// TIA Portal V20 export
ORGANIZATION_BLOCK "T4_Ciclo"   // OB127, LAD, ProgramCycle
TITLE = T4_Ciclo
{ S7_Optimized_Access := 'TRUE' }
AUTHOR : IA
FAMILY : PRUEBA
VERSION : 0.1
// Tanda 1: llama a todas las pruebas
// stored: AutoNumber false, IsIECCheckEnabled false, SetENOAutomatically false
   VAR_INPUT
      Initial_Call : Bool;
      Remanence : Bool;
   END_VAR
BEGIN

REGION Network 1: T4_Base
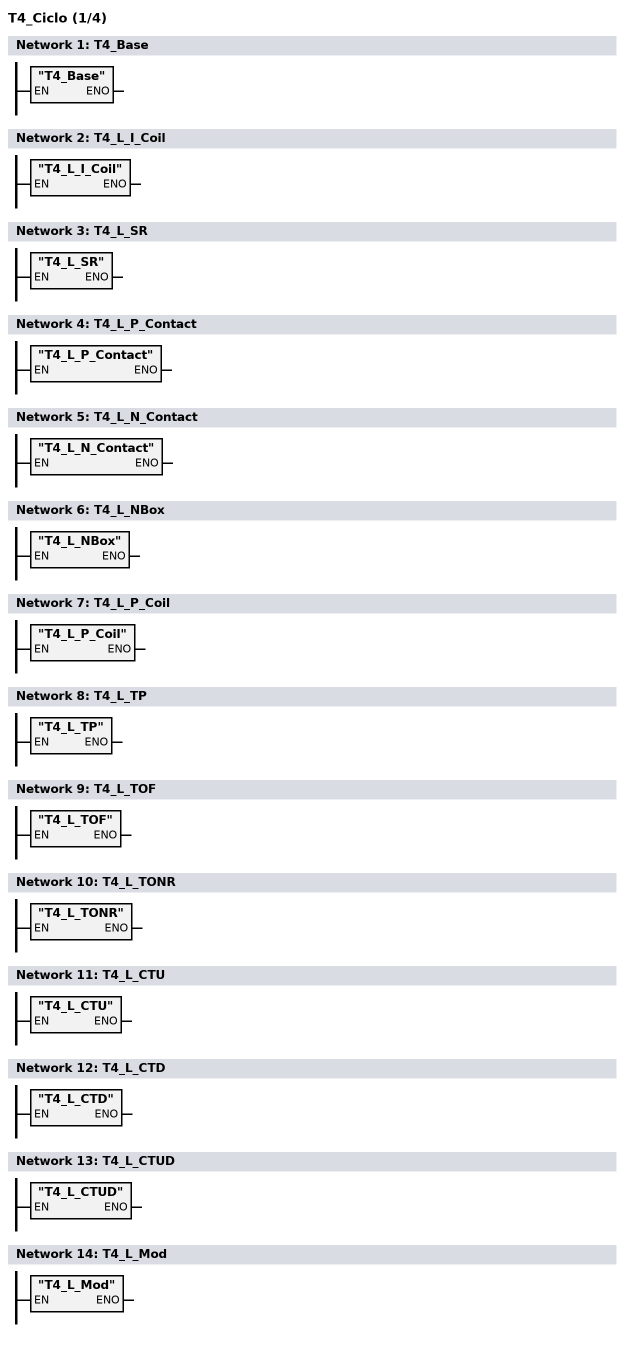
   RUNG wire#powerrail
      "T4_Base"()
   END_RUNG
   // the same network as SCL:
   "T4_Base"();
END_REGION

REGION Network 2: T4_L_I_Coil
   RUNG wire#powerrail
      "T4_L_I_Coil"()
   END_RUNG
   // the same network as SCL:
   "T4_L_I_Coil"();
END_REGION

REGION Network 3: T4_L_SR
   RUNG wire#powerrail
      "T4_L_SR"()
   END_RUNG
   // the same network as SCL:
   "T4_L_SR"();
END_REGION

REGION Network 4: T4_L_P_Contact
   RUNG wire#powerrail
      "T4_L_P_Contact"()
   END_RUNG
   // the same network as SCL:
   "T4_L_P_Contact"();
END_REGION

REGION Network 5: T4_L_N_Contact
   RUNG wire#powerrail
      "T4_L_N_Contact"()
   END_RUNG
   // the same network as SCL:
   "T4_L_N_Contact"();
END_REGION

REGION Network 6: T4_L_NBox
   RUNG wire#powerrail
      "T4_L_NBox"()
   END_RUNG
   // the same network as SCL:
   "T4_L_NBox"();
END_REGION

REGION Network 7: T4_L_P_Coil
   RUNG wire#powerrail
      "T4_L_P_Coil"()
   END_RUNG
   // the same network as SCL:
   "T4_L_P_Coil"();
END_REGION

REGION Network 8: T4_L_TP
   RUNG wire#powerrail
      "T4_L_TP"()
   END_RUNG
   // the same network as SCL:
   "T4_L_TP"();
END_REGION

REGION Network 9: T4_L_TOF
   RUNG wire#powerrail
      "T4_L_TOF"()
   END_RUNG
   // the same network as SCL:
   "T4_L_TOF"();
END_REGION

REGION Network 10: T4_L_TONR
   RUNG wire#powerrail
      "T4_L_TONR"()
   END_RUNG
   // the same network as SCL:
   "T4_L_TONR"();
END_REGION

REGION Network 11: T4_L_CTU
   RUNG wire#powerrail
      "T4_L_CTU"()
   END_RUNG
   // the same network as SCL:
   "T4_L_CTU"();
END_REGION

REGION Network 12: T4_L_CTD
   RUNG wire#powerrail
      "T4_L_CTD"()
   END_RUNG
   // the same network as SCL:
   "T4_L_CTD"();
END_REGION

REGION Network 13: T4_L_CTUD
   RUNG wire#powerrail
      "T4_L_CTUD"()
   END_RUNG
   // the same network as SCL:
   "T4_L_CTUD"();
END_REGION

REGION Network 14: T4_L_Mod
   RUNG wire#powerrail
      "T4_L_Mod"()
   END_RUNG
   // the same network as SCL:
   "T4_L_Mod"();
END_REGION

REGION Network 15: T4_L_Neg
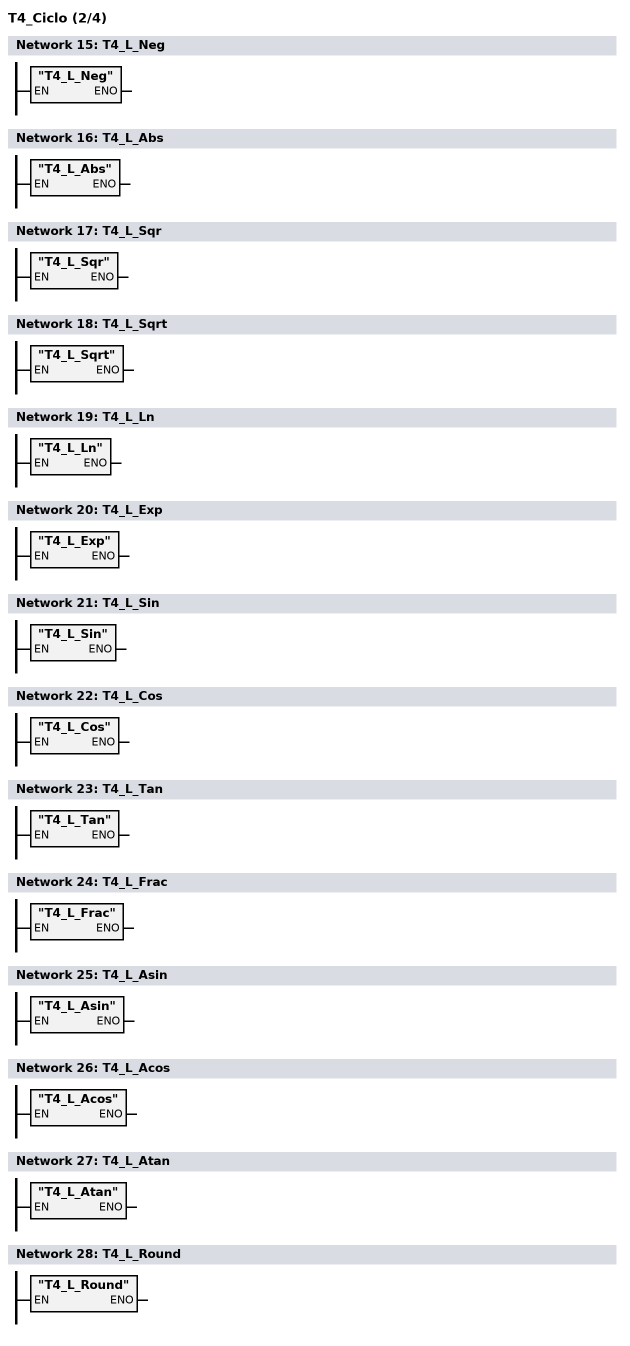
   RUNG wire#powerrail
      "T4_L_Neg"()
   END_RUNG
   // the same network as SCL:
   "T4_L_Neg"();
END_REGION

REGION Network 16: T4_L_Abs
   RUNG wire#powerrail
      "T4_L_Abs"()
   END_RUNG
   // the same network as SCL:
   "T4_L_Abs"();
END_REGION

REGION Network 17: T4_L_Sqr
   RUNG wire#powerrail
      "T4_L_Sqr"()
   END_RUNG
   // the same network as SCL:
   "T4_L_Sqr"();
END_REGION

REGION Network 18: T4_L_Sqrt
   RUNG wire#powerrail
      "T4_L_Sqrt"()
   END_RUNG
   // the same network as SCL:
   "T4_L_Sqrt"();
END_REGION

REGION Network 19: T4_L_Ln
   RUNG wire#powerrail
      "T4_L_Ln"()
   END_RUNG
   // the same network as SCL:
   "T4_L_Ln"();
END_REGION

REGION Network 20: T4_L_Exp
   RUNG wire#powerrail
      "T4_L_Exp"()
   END_RUNG
   // the same network as SCL:
   "T4_L_Exp"();
END_REGION

REGION Network 21: T4_L_Sin
   RUNG wire#powerrail
      "T4_L_Sin"()
   END_RUNG
   // the same network as SCL:
   "T4_L_Sin"();
END_REGION

REGION Network 22: T4_L_Cos
   RUNG wire#powerrail
      "T4_L_Cos"()
   END_RUNG
   // the same network as SCL:
   "T4_L_Cos"();
END_REGION

REGION Network 23: T4_L_Tan
   RUNG wire#powerrail
      "T4_L_Tan"()
   END_RUNG
   // the same network as SCL:
   "T4_L_Tan"();
END_REGION

REGION Network 24: T4_L_Frac
   RUNG wire#powerrail
      "T4_L_Frac"()
   END_RUNG
   // the same network as SCL:
   "T4_L_Frac"();
END_REGION

REGION Network 25: T4_L_Asin
   RUNG wire#powerrail
      "T4_L_Asin"()
   END_RUNG
   // the same network as SCL:
   "T4_L_Asin"();
END_REGION

REGION Network 26: T4_L_Acos
   RUNG wire#powerrail
      "T4_L_Acos"()
   END_RUNG
   // the same network as SCL:
   "T4_L_Acos"();
END_REGION

REGION Network 27: T4_L_Atan
   RUNG wire#powerrail
      "T4_L_Atan"()
   END_RUNG
   // the same network as SCL:
   "T4_L_Atan"();
END_REGION

REGION Network 28: T4_L_Round
   RUNG wire#powerrail
      "T4_L_Round"()
   END_RUNG
   // the same network as SCL:
   "T4_L_Round"();
END_REGION

REGION Network 29: T4_L_Ceil
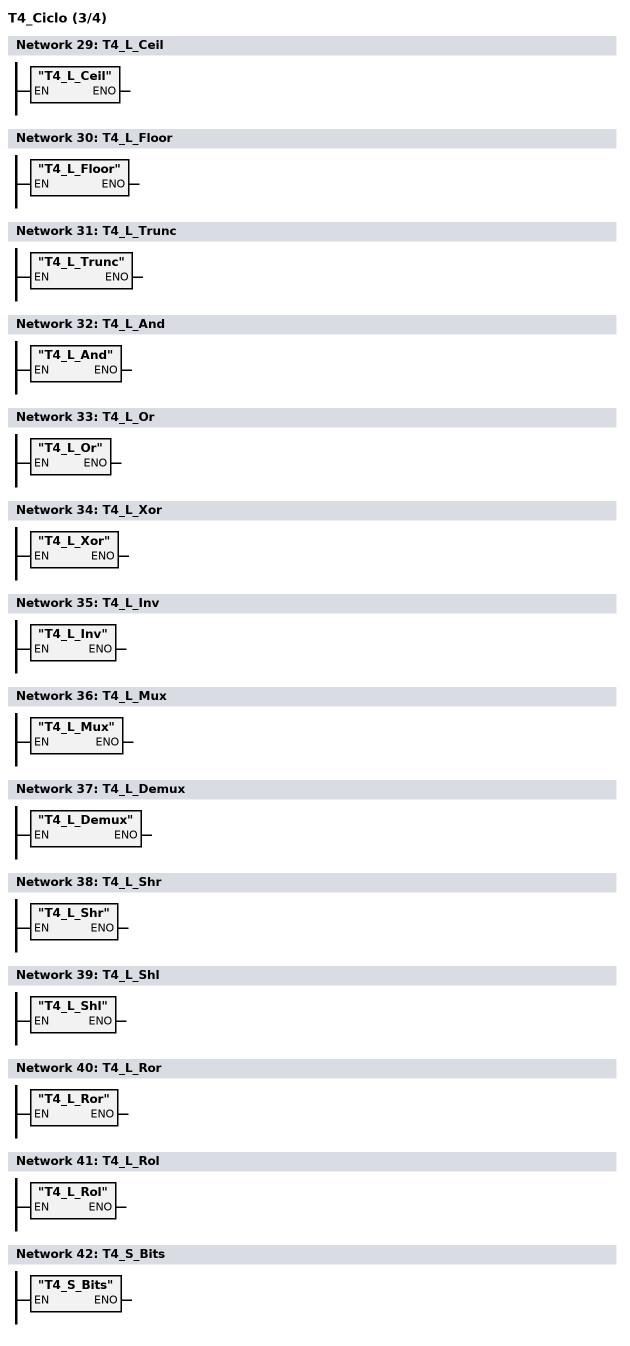
   RUNG wire#powerrail
      "T4_L_Ceil"()
   END_RUNG
   // the same network as SCL:
   "T4_L_Ceil"();
END_REGION

REGION Network 30: T4_L_Floor
   RUNG wire#powerrail
      "T4_L_Floor"()
   END_RUNG
   // the same network as SCL:
   "T4_L_Floor"();
END_REGION

REGION Network 31: T4_L_Trunc
   RUNG wire#powerrail
      "T4_L_Trunc"()
   END_RUNG
   // the same network as SCL:
   "T4_L_Trunc"();
END_REGION

REGION Network 32: T4_L_And
   RUNG wire#powerrail
      "T4_L_And"()
   END_RUNG
   // the same network as SCL:
   "T4_L_And"();
END_REGION

REGION Network 33: T4_L_Or
   RUNG wire#powerrail
      "T4_L_Or"()
   END_RUNG
   // the same network as SCL:
   "T4_L_Or"();
END_REGION

REGION Network 34: T4_L_Xor
   RUNG wire#powerrail
      "T4_L_Xor"()
   END_RUNG
   // the same network as SCL:
   "T4_L_Xor"();
END_REGION

REGION Network 35: T4_L_Inv
   RUNG wire#powerrail
      "T4_L_Inv"()
   END_RUNG
   // the same network as SCL:
   "T4_L_Inv"();
END_REGION

REGION Network 36: T4_L_Mux
   RUNG wire#powerrail
      "T4_L_Mux"()
   END_RUNG
   // the same network as SCL:
   "T4_L_Mux"();
END_REGION

REGION Network 37: T4_L_Demux
   RUNG wire#powerrail
      "T4_L_Demux"()
   END_RUNG
   // the same network as SCL:
   "T4_L_Demux"();
END_REGION

REGION Network 38: T4_L_Shr
   RUNG wire#powerrail
      "T4_L_Shr"()
   END_RUNG
   // the same network as SCL:
   "T4_L_Shr"();
END_REGION

REGION Network 39: T4_L_Shl
   RUNG wire#powerrail
      "T4_L_Shl"()
   END_RUNG
   // the same network as SCL:
   "T4_L_Shl"();
END_REGION

REGION Network 40: T4_L_Ror
   RUNG wire#powerrail
      "T4_L_Ror"()
   END_RUNG
   // the same network as SCL:
   "T4_L_Ror"();
END_REGION

REGION Network 41: T4_L_Rol
   RUNG wire#powerrail
      "T4_L_Rol"()
   END_RUNG
   // the same network as SCL:
   "T4_L_Rol"();
END_REGION

REGION Network 42: T4_S_Bits
   RUNG wire#powerrail
      "T4_S_Bits"()
   END_RUNG
   // the same network as SCL:
   "T4_S_Bits"();
END_REGION

REGION Network 43: T4_S_Tiempo
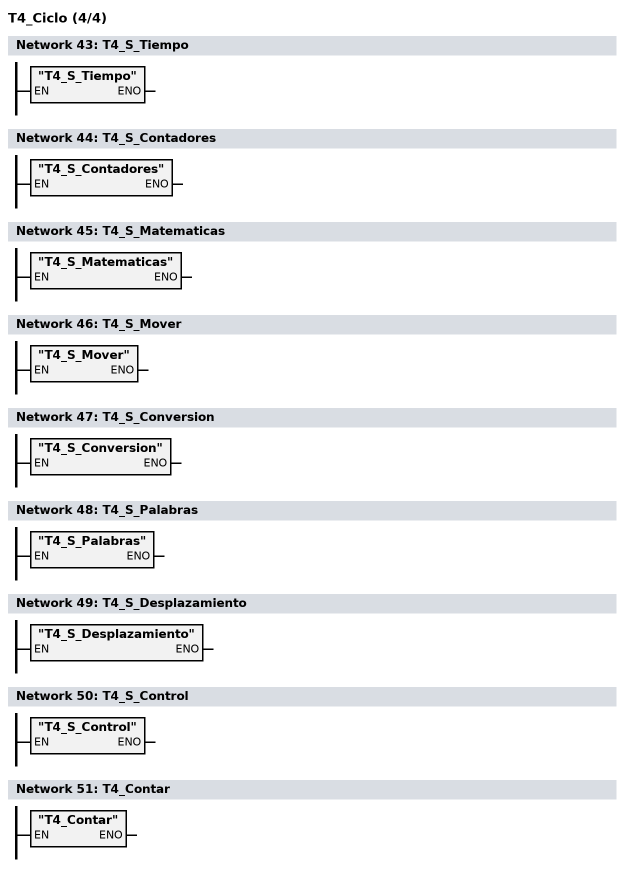
   RUNG wire#powerrail
      "T4_S_Tiempo"()
   END_RUNG
   // the same network as SCL:
   "T4_S_Tiempo"();
END_REGION

REGION Network 44: T4_S_Contadores
   RUNG wire#powerrail
      "T4_S_Contadores"()
   END_RUNG
   // the same network as SCL:
   "T4_S_Contadores"();
END_REGION

REGION Network 45: T4_S_Matematicas
   RUNG wire#powerrail
      "T4_S_Matematicas"()
   END_RUNG
   // the same network as SCL:
   "T4_S_Matematicas"();
END_REGION

REGION Network 46: T4_S_Mover
   RUNG wire#powerrail
      "T4_S_Mover"()
   END_RUNG
   // the same network as SCL:
   "T4_S_Mover"();
END_REGION

REGION Network 47: T4_S_Conversion
   RUNG wire#powerrail
      "T4_S_Conversion"()
   END_RUNG
   // the same network as SCL:
   "T4_S_Conversion"();
END_REGION

REGION Network 48: T4_S_Palabras
   RUNG wire#powerrail
      "T4_S_Palabras"()
   END_RUNG
   // the same network as SCL:
   "T4_S_Palabras"();
END_REGION

REGION Network 49: T4_S_Desplazamiento
   RUNG wire#powerrail
      "T4_S_Desplazamiento"()
   END_RUNG
   // the same network as SCL:
   "T4_S_Desplazamiento"();
END_REGION

REGION Network 50: T4_S_Control
   RUNG wire#powerrail
      "T4_S_Control"()
   END_RUNG
   // the same network as SCL:
   "T4_S_Control"();
END_REGION

REGION Network 51: T4_Contar
   RUNG wire#powerrail
      "T4_Contar"()
   END_RUNG
   // the same network as SCL:
   "T4_Contar"();
END_REGION
END_ORGANIZATION_BLOCK
